FUNCTION_BLOCK "FB_Station"
TITLE = 'Mixing station: devices, sequence, interlocks, alarms, line interface'
{ S7_Optimized_Access := 'TRUE' }
AUTHOR : Demo
VERSION : 0.1
   VAR
      LT101 : "FB_AnalogIn";   // Tank level transmitter, 0..100 %
      TT301 : "FB_AnalogIn";   // Tank temperature transmitter, 0..120 degC
      XV101 : "FB_Valve";   // Inlet valve ingredient A
      XV102 : "FB_Valve";   // Inlet valve ingredient B
      M201 : "FB_VFD";   // Agitator on a VFD
      P401 : "FB_Motor";   // Outlet pump
      Alarms : "FB_AlarmHandler";   // Latches alarm conditions into DB_Alarms
      tMesHb {InstructionName := 'TON_TIME'; LibVersion := '1.0'} : TON_TIME;   // MES heartbeat watchdog (5 s)
      tOwnHb {InstructionName := 'TON_TIME'; LibVersion := '1.0'} : TON_TIME;   // 1 s pulse for our own heartbeat
      OwnHbDone : Bool;   // TRUE for one cycle after each 1 s pulse
      LastMesHb : Int;   // MES heartbeat value in the previous cycle
      tHeat {InstructionName := 'TON_TIME'; LibVersion := '1.0'} : TON_TIME;   // Heater on without a break (60 s)
      TempAtHeatOn : Real;   // Temperature when the heater last switched on [degC]
      NoHeating : Bool;   // Heater on for 60 s but temperature rose less than 2 degC
   END_VAR

BEGIN
	// ---------- Analog inputs ----------
	#LT101(Raw := "DB_IO".LT101_Raw, RangeLo := 0.0, RangeHi := 100.0, LimitHigh := 95.0, LimitLow := 5.0);
	#TT301(Raw := "DB_IO".TT301_Raw, RangeLo := 0.0, RangeHi := 120.0, LimitHigh := 90.0, LimitLow := 0.0);

	// ---------- Sequence ----------
	// Own instance DB, not a multi-instance: GRAPH blocks (plc-demo/graph) cannot be multi-instances.
	"DB_BatchSequence"(Start := "DB_IO".PB_Start OR "DB_LineInterface".MES_StartRequest,
	                   Stop := "DB_IO".PB_Stop,
	                   Auto := "DB_IO".SW_Auto,
	                   AnyFault := "DB_Alarms".AnyFault,
	                   EStopOK := "DB_IO".EStop_OK,
	                   Level := #LT101.Value,
	                   Temp := #TT301.Value,
	                   FillerReady := "DB_LineInterface".Filler_ReadyToReceive);

	// ---------- Devices with interlocks ----------
	// Inlet valves may not open when the level is high (overflow protection)
	#XV101(Open := "DB_BatchSequence".OpenXV101, Permit := NOT #LT101.High AND NOT #LT101.WireBreak,
	       ZSO := "DB_IO".XV101_ZSO, ZSC := "DB_IO".XV101_ZSC);
	#XV102(Open := "DB_BatchSequence".OpenXV102, Permit := NOT #LT101.High AND NOT #LT101.WireBreak,
	       ZSO := "DB_IO".XV102_ZSO, ZSC := "DB_IO".XV102_ZSC);
	"DB_IO".XV101_OpenCmd := #XV101.Out;
	"DB_IO".XV102_OpenCmd := #XV102.Out;

	// Agitator may only run with the blades covered (level above 20 %)
	#M201(Run := "DB_BatchSequence".RunM201, Permit := #LT101.Value > 20.0 AND "DB_IO".EStop_OK,
	      SpeedSP := "DB_BatchSequence".SpeedM201, SpeedPV := "DB_IO".M201_SpeedPV,
	      Ready := "DB_IO".M201_DriveReady, DriveFault := "DB_IO".M201_DriveFault);
	"DB_IO".M201_RunCmd := #M201.RunOut;
	"DB_IO".M201_SpeedSP := #M201.SpeedOut;

	// Heater only with the agitator running (no local overheating) and no overtemperature
	"DB_IO".E301_OnCmd := "DB_BatchSequence".HeatE301 AND #M201.AtSpeed AND NOT "DB_IO".E301_OverTemp AND NOT #TT301.WireBreak;

	// Heating check: heater on for 60 s without a break but the temperature rose less than 2 degC.
	// The window starts again each time the heater switches on, also after a halt.
	IF NOT "DB_IO".E301_OnCmd THEN
	    #TempAtHeatOn := #TT301.Value;
	END_IF;
	#tHeat(IN := "DB_IO".E301_OnCmd, PT := T#60S);
	#NoHeating := #tHeat.Q AND #TT301.Value < #TempAtHeatOn + 2.0;

	// Pump may not run dry
	#P401(Run := "DB_BatchSequence".RunP401, Permit := #LT101.Value > 0.5 AND "DB_IO".EStop_OK,
	      RunFb := "DB_IO".P401_RunFb, Trip := "DB_IO".P401_MotorTrip);
	"DB_IO".P401_RunCmd := #P401.Out;

	// ---------- Line interface (data exchange) ----------
	#tMesHb(IN := "DB_LineInterface".MES_Heartbeat = #LastMesHb, PT := T#5S);
	#LastMesHb := "DB_LineInterface".MES_Heartbeat;
	#tOwnHb(IN := NOT #OwnHbDone, PT := T#1S);
	#OwnHbDone := #tOwnHb.Q;
	IF #OwnHbDone THEN
	    "DB_LineInterface".Station_Heartbeat := ("DB_LineInterface".Station_Heartbeat + 1) MOD 30000;
	END_IF;
	IF "DB_BatchSequence".Step = 0 THEN
	    "DB_Recipe".RecipeNo := "DB_LineInterface".MES_RecipeNo;
	END_IF;
	"DB_LineInterface".Station_Running := "DB_BatchSequence".Running;
	"DB_LineInterface".Station_Draining := "DB_BatchSequence".Step = 50;
	"DB_LineInterface".Batch_Done := "DB_BatchSequence".BatchDone;
	IF "DB_BatchSequence".BatchDone THEN
	    "DB_LineInterface".Batch_Count := "DB_LineInterface".Batch_Count + 1;
	END_IF;

	// ---------- Alarms ----------
	#Alarms(Reset := "DB_IO".PB_Reset,
	        EStop := NOT "DB_IO".EStop_OK,
	        XV101_NotOpen := #XV101.FaultNotOpen,
	        XV101_NotClosed := #XV101.FaultNotClosed,
	        XV102_NotOpen := #XV102.FaultNotOpen,
	        XV102_NotClosed := #XV102.FaultNotClosed,
	        M201_DriveFault := #M201.FaultDrive,
	        M201_SpeedDev := #M201.FaultSpeedDev,
	        M201_NotReady := #M201.NotReady,
	        E301_OverTemp := "DB_IO".E301_OverTemp,
	        P401_Trip := #P401.FaultTrip,
	        P401_NoFeedback := #P401.FaultNoFeedback,
	        LT101_WireBreak := #LT101.WireBreak,
	        LT101_HighHigh := #LT101.High,
	        TT301_WireBreak := #TT301.WireBreak,
	        TT301_High := #TT301.High,
	        Step10_Timeout := "DB_BatchSequence".TimeoutStep10,
	        Step20_Timeout := "DB_BatchSequence".TimeoutStep20,
	        Step30_Timeout := "DB_BatchSequence".TimeoutStep30,
	        Step50_Timeout := "DB_BatchSequence".TimeoutStep50,
	        E301_NoHeating := #NoHeating,
	        Filler_NotReady := "DB_BatchSequence".WaitFillerTooLong,
	        MES_HeartbeatLost := #tMesHb.Q,
	        RecipeInvalid := "DB_BatchSequence".StartRecipeInvalid,
	        NotInAuto := "DB_BatchSequence".StartNotAuto,
	        TankNotEmpty := "DB_BatchSequence".StartTankNotEmpty);
END_FUNCTION_BLOCK
